Fanuc KAREL source: IO0191.KL

PROGRAM IO0191
%NOLOCKGROUP
ROUTINE RTEST
VAR
  I : INTEGER
  STATUS : INTEGER
  ENTRY : INTEGER
  A : ARRAY[3] OF INTEGER
  B : BOOLEAN
  R : REAL
  P : XYZWPR
  JPOS : JOINTPOS
  PF : POSITION
BEGIN
  I = 1
  A[1] = 2
  B = TRUE
  R = 1.0
  WAIT FOR DIN[A[I]] = ON
END RTEST
BEGIN
  RTEST
END IO0191
